  movel([-0.141321, -0.804315, -2.796072, -1.112001, 1.570796, 1.429476],accel_mss,speed_ms,0,blend_radius_m)
  movel([-0.146733, -0.812986, -2.794574, -1.104829, 1.570796, 1.424064],accel_mss,speed_ms,0,blend_radius_m)
  movel([-0.151447, -0.821414, -2.793080, -1.097895, 1.570796, 1.419350],accel_mss,speed_ms,0,blend_radius_m)
  movel([-0.155435, -0.829598, -2.791592, -1.091199, 1.570796, 1.415362],accel_mss,speed_ms,0,blend_radius_m)
  movel([-0.157149, -0.833600, -2.790851, -1.087938, 1.570796, 1.413648],accel_mss,speed_ms,0,blend_radius_m)
  movel([-0.159989, -0.841407, -2.789381, -1.081601, 1.570796, 1.410807],accel_mss,speed_ms,0,blend_radius_m)
  movel([-0.161109, -0.845218, -2.788651, -1.078520, 1.570796, 1.409688],accel_mss,speed_ms,0,blend_radius_m)
  movel([-0.162732, -0.852643, -2.787205, -1.072541, 1.570796, 1.408064],accel_mss,speed_ms,0,blend_radius_m)
  movel([-0.163230, -0.856264, -2.786488, -1.069637, 1.570796, 1.407566],accel_mss,speed_ms,0,blend_radius_m)
  movel([-0.163513, -0.859817, -2.785778, -1.066794, 1.570796, 1.407283],accel_mss,speed_ms,0,blend_radius_m)
  movel([-0.163602, -0.864722, -2.784786, -1.062881, 1.570796, 1.407194],accel_mss,speed_ms,0,blend_radius_m)
  movel([-0.163380, -0.869441, -2.783818, -1.059131, 1.570796, 1.407417],accel_mss,speed_ms,0,blend_radius_m)
  movel([-0.162870, -0.873957, -2.782879, -1.055553, 1.570796, 1.407926],accel_mss,speed_ms,0,blend_radius_m)
  movel([-0.162104, -0.878276, -2.781970, -1.052143, 1.570796, 1.408692],accel_mss,speed_ms,0,blend_radius_m)
  movel([-0.161097, -0.882370, -2.781098, -1.048921, 1.570796, 1.409700],accel_mss,speed_ms,0,blend_radius_m)
  movel([-0.159870, -0.886230, -2.780267, -1.045892, 1.570796, 1.410927],accel_mss,speed_ms,0,blend_radius_m)
  movel([-0.158448, -0.889851, -2.779479, -1.043059, 1.570796, 1.412348],accel_mss,speed_ms,0,blend_radius_m)
  movel([-0.156848, -0.893214, -2.778740, -1.040435, 1.570796, 1.413948],accel_mss,speed_ms,0,blend_radius_m)
  movel([-0.149158, -0.904985, -2.776098, -1.031305, 1.570796, 1.421638],accel_mss,speed_ms,0,blend_radius_m)
  movel([-0.143209, -0.914586, -2.773880, -1.023923, 1.570796, 1.427587],accel_mss,speed_ms,0,blend_radius_m)
  movel([-0.142775, -0.915615, -2.773639, -1.023135, 1.570796, 1.428021],accel_mss,speed_ms,0,blend_radius_m)
  movel([-0.135600, -0.906199, -2.775821, -1.030369, 1.570796, 1.435197],accel_mss,speed_ms,0,blend_radius_m)
  movel([-0.127938, -0.896903, -2.777921, -1.037564, 1.570796, 1.442859],accel_mss,speed_ms,0,blend_radius_m)
  movel([-0.119839, -0.887763, -2.779934, -1.044692, 1.570796, 1.450957],accel_mss,speed_ms,0,blend_radius_m)
  movel([-0.111369, -0.878821, -2.781854, -1.051713, 1.570796, 1.459427],accel_mss,speed_ms,0,blend_radius_m)
  movel([-0.102591, -0.870130, -2.783675, -1.058584, 1.570796, 1.468205],accel_mss,speed_ms,0,blend_radius_m)
  movel([-0.093574, -0.861730, -2.785393, -1.065267, 1.570796, 1.477222],accel_mss,speed_ms,0,blend_radius_m)
  movel([-0.084386, -0.853674, -2.787002, -1.071713, 1.570796, 1.486410],accel_mss,speed_ms,0,blend_radius_m)
  movel([-0.075105, -0.846013, -2.788497, -1.077879, 1.570796, 1.495692],accel_mss,speed_ms,0,blend_radius_m)
  movel([-0.070692, -0.842600, -2.789153, -1.080635, 1.570796, 1.500104],accel_mss,speed_ms,0,blend_radius_m)
  movel([-0.066171, -0.839349, -2.789772, -1.083268, 1.570796, 1.504626],accel_mss,speed_ms,0,blend_radius_m)
  movel([-0.061579, -0.836295, -2.790347, -1.085746, 1.570796, 1.509218],accel_mss,speed_ms,0,blend_radius_m)
  movel([-0.056967, -0.833486, -2.790873, -1.088031, 1.570796, 1.513830],accel_mss,speed_ms,0,blend_radius_m)
  movel([-0.052375, -0.830958, -2.791341, -1.090090, 1.570796, 1.518421],accel_mss,speed_ms,0,blend_radius_m)
  movel([-0.047846, -0.828755, -2.791747, -1.091887, 1.570796, 1.522951],accel_mss,speed_ms,0,blend_radius_m)
  movel([-0.043425, -0.826913, -2.792084, -1.093392, 1.570796, 1.527371],accel_mss,speed_ms,0,blend_radius_m)
  movel([-0.039161, -0.825474, -2.792346, -1.094569, 1.570796, 1.531636],accel_mss,speed_ms,0,blend_radius_m)
  movel([-0.035094, -0.824478, -2.792527, -1.095384, 1.570796, 1.535702],accel_mss,speed_ms,0,blend_radius_m)
  movel([-0.031268, -0.823960, -2.792621, -1.095808, 1.570796, 1.539528],accel_mss,speed_ms,0,blend_radius_m)
  movel([-0.027734, -0.823963, -2.792620, -1.095806, 1.570796, 1.543062],accel_mss,speed_ms,0,blend_radius_m)
  movel([-0.024533, -0.824519, -2.792520, -1.095350, 1.570796, 1.546264],accel_mss,speed_ms,0,blend_radius_m)
  movel([-0.021709, -0.825663, -2.792312, -1.094414, 1.570796, 1.549087],accel_mss,speed_ms,0,blend_radius_m)
  movel([-0.019297, -0.827423, -2.791991, -1.092975, 1.570796, 1.551499],accel_mss,speed_ms,0,blend_radius_m)
  movel([-0.017345, -0.829831, -2.791549, -1.091009, 1.570796, 1.553452],accel_mss,speed_ms,0,blend_radius_m)
  movel([-0.015891, -0.832916, -2.790978, -1.088494, 1.570796, 1.554905],accel_mss,speed_ms,0,blend_radius_m)
  movel([-0.014708, -0.837711, -2.790081, -1.084597, 1.570796, 1.556088],accel_mss,speed_ms,0,blend_radius_m)
  movel([-0.014174, -0.843160, -2.789046, -1.080183, 1.570796, 1.556622],accel_mss,speed_ms,0,blend_radius_m)
  movel([-0.014196, -0.849111, -2.787897, -1.075382, 1.570796, 1.556600],accel_mss,speed_ms,0,blend_radius_m)
  movel([-0.014673, -0.855417, -2.786657, -1.070315, 1.570796, 1.556123],accel_mss,speed_ms,0,blend_radius_m)
  movel([-0.015515, -0.861935, -2.785351, -1.065103, 1.570796, 1.555282],accel_mss,speed_ms,0,blend_radius_m)
  movel([-0.016634, -0.868531, -2.784005, -1.059853, 1.570796, 1.554162],accel_mss,speed_ms,0,blend_radius_m)
  movel([-0.019330, -0.881416, -2.781302, -1.049671, 1.570796, 1.551466],accel_mss,speed_ms,0,blend_radius_m)
  movel([-0.021385, -0.889588, -2.779536, -1.043265, 1.570796, 1.549411],accel_mss,speed_ms,0,blend_radius_m)
  movel([-0.023782, -0.897714, -2.777740, -1.036935, 1.570796, 1.547015],accel_mss,speed_ms,0,blend_radius_m)
  movel([-0.026474, -0.905794, -2.775914, -1.030681, 1.570796, 1.544323],accel_mss,speed_ms,0,blend_radius_m)
  movel([-0.029419, -0.913847, -2.774053, -1.024489, 1.570796, 1.541377],accel_mss,speed_ms,0,blend_radius_m)
  movel([-0.032573, -0.921870, -2.772158, -1.018361, 1.570796, 1.538223],accel_mss,speed_ms,0,blend_radius_m)
  movel([-0.035892, -0.929878, -2.770225, -1.012287, 1.570796, 1.534904],accel_mss,speed_ms,0,blend_radius_m)
  movel([-0.042880, -0.945892, -2.766232, -1.000265, 1.570796, 1.527916],accel_mss,speed_ms,0,blend_radius_m)
  movel([-0.036325, -0.946186, -2.766157, -1.000046, 1.570796, 1.534471],accel_mss,speed_ms,0,blend_radius_m)
  movel([-0.032953, -0.946594, -2.766053, -0.999742, 1.570796, 1.537843],accel_mss,speed_ms,0,blend_radius_m)
  movel([-0.030089, -0.947502, -2.765821, -0.999065, 1.570796, 1.540707],accel_mss,speed_ms,0,blend_radius_m)
  movel([-0.028984, -0.948223, -2.765637, -0.998529, 1.570796, 1.541813],accel_mss,speed_ms,0,blend_radius_m)
  movel([-0.028168, -0.949162, -2.765396, -0.997831, 1.570796, 1.542628],accel_mss,speed_ms,0,blend_radius_m)
  movel([-0.027690, -0.950344, -2.765092, -0.996953, 1.570796, 1.543106],accel_mss,speed_ms,0,blend_radius_m)
  movel([-0.027603, -0.951798, -2.764716, -0.995875, 1.570796, 1.543193],accel_mss,speed_ms,0,blend_radius_m)
  movel([-0.027958, -0.953548, -2.764263, -0.994579, 1.570796, 1.542838],accel_mss,speed_ms,0,blend_radius_m)
  movel([-0.028810, -0.955631, -2.763720, -0.993039, 1.570796, 1.541986],accel_mss,speed_ms,0,blend_radius_m)
  movel([-0.030204, -0.958070, -2.763080, -0.991239, 1.570796, 1.540592],accel_mss,speed_ms,0,blend_radius_m)
  movel([-0.032189, -0.960886, -2.762337, -0.989166, 1.570796, 1.538607],accel_mss,speed_ms,0,blend_radius_m)
  movel([-0.034030, -0.963178, -2.761728, -0.987484, 1.570796, 1.536766],accel_mss,speed_ms,0,blend_radius_m)
  movel([-0.035882, -0.965239, -2.761177, -0.985973, 1.570796, 1.534914],accel_mss,speed_ms,0,blend_radius_m)
  movel([-0.037742, -0.967088, -2.760680, -0.984621, 1.570796, 1.533055],accel_mss,speed_ms,0,blend_radius_m)
  movel([-0.041487, -0.970225, -2.759832, -0.982332, 1.570796, 1.529310],accel_mss,speed_ms,0,blend_radius_m)
  movel([-0.043369, -0.971550, -2.759471, -0.981368, 1.570796, 1.527427],accel_mss,speed_ms,0,blend_radius_m)
  movel([-0.047159, -0.973809, -2.758854, -0.979726, 1.570796, 1.523638],accel_mss,speed_ms,0,blend_radius_m)
  movel([-0.050963, -0.975658, -2.758346, -0.978385, 1.570796, 1.519833],accel_mss,speed_ms,0,blend_radius_m)
  movel([-0.054779, -0.977239, -2.757910, -0.977241, 1.570796, 1.516017],accel_mss,speed_ms,0,blend_radius_m)
  movel([-0.062394, -0.980130, -2.757107, -0.975152, 1.570796, 1.508402],accel_mss,speed_ms,0,blend_radius_m)
  movel([-0.066370, -0.986523, -2.755311, -0.970555, 1.570796, 1.504426],accel_mss,speed_ms,0,blend_radius_m)
  movel([-0.068546, -0.989715, -2.754403, -0.968271, 1.570796, 1.502250],accel_mss,speed_ms,0,blend_radius_m)
  movel([-0.070857, -0.992817, -2.753513, -0.966058, 1.570796, 1.499939],accel_mss,speed_ms,0,blend_radius_m)
  movel([-0.073309, -0.995761, -2.752662, -0.963965, 1.570796, 1.497488],accel_mss,speed_ms,0,blend_radius_m)
  movel([-0.075903, -0.998481, -2.751871, -0.962038, 1.570796, 1.494894],accel_mss,speed_ms,0,blend_radius_m)
  movel([-0.078648, -1.000910, -2.751159, -0.960321, 1.570796, 1.492149],accel_mss,speed_ms,0,blend_radius_m)
  movel([-0.081555, -1.002990, -2.750546, -0.958854, 1.570796, 1.489241],accel_mss,speed_ms,0,blend_radius_m)
  movel([-0.083598, -1.004037, -2.750236, -0.958116, 1.570796, 1.487198],accel_mss,speed_ms,0,blend_radius_m)
  movel([-0.085214, -1.004394, -2.750130, -0.957865, 1.570796, 1.485582],accel_mss,speed_ms,0,blend_radius_m)
  movel([-0.086450, -1.004162, -2.750199, -0.958028, 1.570796, 1.484347],accel_mss,speed_ms,0,blend_radius_m)
  movel([-0.087346, -1.003436, -2.750414, -0.958539, 1.570796, 1.483451],accel_mss,speed_ms,0,blend_radius_m)
  movel([-0.087946, -1.002312, -2.750746, -0.959331, 1.570796, 1.482851],accel_mss,speed_ms,0,blend_radius_m)
  movel([-0.088287, -1.000895, -2.751163, -0.960331, 1.570796, 1.482509],accel_mss,speed_ms,0,blend_radius_m)
  movel([-0.088418, -0.999280, -2.751637, -0.961472, 1.570796, 1.482378],accel_mss,speed_ms,0,blend_radius_m)
  movel([-0.088369, -0.997561, -2.752139, -0.962689, 1.570796, 1.482428],accel_mss,speed_ms,0,blend_radius_m)
  movel([-0.087893, -0.993747, -2.753245, -0.965397, 1.570796, 1.482904],accel_mss,speed_ms,0,blend_radius_m)
  movel([-0.087059, -0.989798, -2.754379, -0.968212, 1.570796, 1.483737],accel_mss,speed_ms,0,blend_radius_m)
  movel([-0.084858, -0.981561, -2.756707, -0.974120, 1.570796, 1.485939],accel_mss,speed_ms,0,blend_radius_m)
  movel([-0.093540, -0.980140, -2.757104, -0.975145, 1.570796, 1.477256],accel_mss,speed_ms,0,blend_radius_m)
  movel([-0.102455, -0.979099, -2.757394, -0.975896, 1.570796, 1.468341],accel_mss,speed_ms,0,blend_radius_m)
  movel([-0.111365, -0.978026, -2.757692, -0.976671, 1.570796, 1.459431],accel_mss,speed_ms,0,blend_radius_m)
  movel([-0.115747, -0.977350, -2.757879, -0.977161, 1.570796, 1.455049],accel_mss,speed_ms,0,blend_radius_m)
  movel([-0.120046, -0.976509, -2.758111, -0.977769, 1.570796, 1.450750],accel_mss,speed_ms,0,blend_radius_m)
  movel([-0.124039, -0.975495, -2.758391, -0.978503, 1.570796, 1.446757],accel_mss,speed_ms,0,blend_radius_m)
  movel([-0.127889, -0.974301, -2.758719, -0.979369, 1.570796, 1.442907],accel_mss,speed_ms,0,blend_radius_m)
  movel([-0.135327, -0.971570, -2.759466, -0.981353, 1.570796, 1.435469],accel_mss,speed_ms,0,blend_radius_m)
  movel([-0.142709, -0.968772, -2.760225, -0.983392, 1.570796, 1.428087],accel_mss,speed_ms,0,blend_radius_m)
  movel([-0.150371, -0.966361, -2.760875, -0.985152, 1.570796, 1.420425],accel_mss,speed_ms,0,blend_radius_m)
  movel([-0.152086, -0.971127, -2.759586, -0.981675, 1.570796, 1.418710],accel_mss,speed_ms,0,blend_radius_m)
  movel([-0.153549, -0.975769, -2.758315, -0.978305, 1.570796, 1.417247],accel_mss,speed_ms,0,blend_radius_m)
  movel([-0.154762, -0.980277, -2.757066, -0.975046, 1.570796, 1.416035],accel_mss,speed_ms,0,blend_radius_m)
  movel([-0.155729, -0.984644, -2.755842, -0.971903, 1.570796, 1.415067],accel_mss,speed_ms,0,blend_radius_m)
  movel([-0.156451, -0.988870, -2.754644, -0.968875, 1.570796, 1.414345],accel_mss,speed_ms,0,blend_radius_m)
  movel([-0.156938, -0.992946, -2.753476, -0.965967, 1.570796, 1.413859],accel_mss,speed_ms,0,blend_radius_m)
  movel([-0.157185, -0.996868, -2.752341, -0.963180, 1.570796, 1.413612],accel_mss,speed_ms,0,blend_radius_m)
  movel([-0.157205, -1.000637, -2.751239, -0.960513, 1.570796, 1.413592],accel_mss,speed_ms,0,blend_radius_m)
  movel([-0.156995, -1.004243, -2.750175, -0.957972, 1.570796, 1.413802],accel_mss,speed_ms,0,blend_radius_m)
  movel([-0.156554, -1.007678, -2.749152, -0.955559, 1.570796, 1.414242],accel_mss,speed_ms,0,blend_radius_m)
  movel([-0.155895, -1.010950, -2.748169, -0.953270, 1.570796, 1.414901],accel_mss,speed_ms,0,blend_radius_m)
  movel([-0.155018, -1.014046, -2.747232, -0.951112, 1.570796, 1.415778],accel_mss,speed_ms,0,blend_radius_m)
  movel([-0.153919, -1.016958, -2.746343, -0.949088, 1.570796, 1.416877],accel_mss,speed_ms,0,blend_radius_m)
  movel([-0.152607, -1.019693, -2.745503, -0.947193, 1.570796, 1.418189],accel_mss,speed_ms,0,blend_radius_m)
  movel([-0.151084, -1.022240, -2.744715, -0.945434, 1.570796, 1.419713],accel_mss,speed_ms,0,blend_radius_m)
  movel([-0.149346, -1.024596, -2.743981, -0.943812, 1.570796, 1.421450],accel_mss,speed_ms,0,blend_radius_m)
  movel([-0.146282, -1.027856, -2.742959, -0.941574, 1.570796, 1.424514],accel_mss,speed_ms,0,blend_radius_m)
  movel([-0.142850, -1.030642, -2.742079, -0.939668, 1.570796, 1.427946],accel_mss,speed_ms,0,blend_radius_m)
  movel([-0.139097, -1.033005, -2.741328, -0.938057, 1.570796, 1.431699],accel_mss,speed_ms,0,blend_radius_m)
  movel([-0.135055, -1.034984, -2.740695, -0.936710, 1.570796, 1.435741],accel_mss,speed_ms,0,blend_radius_m)
  movel([-0.130770, -1.036629, -2.740167, -0.935593, 1.570796, 1.440026],accel_mss,speed_ms,0,blend_radius_m)
  movel([-0.126280, -1.037978, -2.739732, -0.934679, 1.570796, 1.444516],accel_mss,speed_ms,0,blend_radius_m)
  movel([-0.121626, -1.039078, -2.739376, -0.933935, 1.570796, 1.449171],accel_mss,speed_ms,0,blend_radius_m)
  movel([-0.116838, -1.039956, -2.739092, -0.933342, 1.570796, 1.453958],accel_mss,speed_ms,0,blend_radius_m)
  movel([-0.106974, -1.041285, -2.738660, -0.932445, 1.570796, 1.463822],accel_mss,speed_ms,0,blend_radius_m)
  movel([-0.096981, -1.042372, -2.738305, -0.931712, 1.570796, 1.473815],accel_mss,speed_ms,0,blend_radius_m)
  movel([-0.089406, -1.043472, -2.737946, -0.930972, 1.570796, 1.481391],accel_mss,speed_ms,0,blend_radius_m)
  movel([-0.086797, -1.043644, -2.737889, -0.930856, 1.570796, 1.484000],accel_mss,speed_ms,0,blend_radius_m)
  movel([-0.082087, -1.043552, -2.737919, -0.930918, 1.570796, 1.488709],accel_mss,speed_ms,0,blend_radius_m)
  movel([-0.081105, -1.043729, -2.737861, -0.930799, 1.570796, 1.489692],accel_mss,speed_ms,0,blend_radius_m)
  movel([-0.080223, -1.044102, -2.737739, -0.930548, 1.570796, 1.490574],accel_mss,speed_ms,0,blend_radius_m)
  movel([-0.079458, -1.044736, -2.737531, -0.930122, 1.570796, 1.491338],accel_mss,speed_ms,0,blend_radius_m)
  movel([-0.078830, -1.045693, -2.737216, -0.929480, 1.570796, 1.491966],accel_mss,speed_ms,0,blend_radius_m)
  movel([-0.078371, -1.047037, -2.736773, -0.928579, 1.570796, 1.492426],accel_mss,speed_ms,0,blend_radius_m)
  movel([-0.078211, -1.048560, -2.736269, -0.927560, 1.570796, 1.492585],accel_mss,speed_ms,0,blend_radius_m)
  movel([-0.078322, -1.050228, -2.735715, -0.926446, 1.570796, 1.492474],accel_mss,speed_ms,0,blend_radius_m)
  movel([-0.078680, -1.052026, -2.735115, -0.925248, 1.570796, 1.492116],accel_mss,speed_ms,0,blend_radius_m)
  movel([-0.079260, -1.053920, -2.734480, -0.923989, 1.570796, 1.491536],accel_mss,speed_ms,0,blend_radius_m)
  movel([-0.080989, -1.057919, -2.733129, -0.921340, 1.570796, 1.489808],accel_mss,speed_ms,0,blend_radius_m)
  movel([-0.082090, -1.059975, -2.732430, -0.919984, 1.570796, 1.488706],accel_mss,speed_ms,0,blend_radius_m)
  movel([-0.084632, -1.064080, -2.731023, -0.917287, 1.570796, 1.486165],accel_mss,speed_ms,0,blend_radius_m)
  movel([-0.087485, -1.068033, -2.729654, -0.914703, 1.570796, 1.483311],accel_mss,speed_ms,0,blend_radius_m)
  movel([-0.090454, -1.071655, -2.728388, -0.912347, 1.570796, 1.480342],accel_mss,speed_ms,0,blend_radius_m)
  movel([-0.093367, -1.074779, -2.727286, -0.910323, 1.570796, 1.477429],accel_mss,speed_ms,0,blend_radius_m)
  movel([-0.097927, -1.079003, -2.725784, -0.907602, 1.570796, 1.472870],accel_mss,speed_ms,0,blend_radius_m)
  movel([-0.100289, -1.080959, -2.725083, -0.906347, 1.570796, 1.470507],accel_mss,speed_ms,0,blend_radius_m)
  movel([-0.102689, -1.082800, -2.724421, -0.905168, 1.570796, 1.468107],accel_mss,speed_ms,0,blend_radius_m)
  movel([-0.107574, -1.086135, -2.723212, -0.903042, 1.570796, 1.463222],accel_mss,speed_ms,0,blend_radius_m)
  movel([-0.112504, -1.088976, -2.722175, -0.901238, 1.570796, 1.458292],accel_mss,speed_ms,0,blend_radius_m)
  movel([-0.117406, -1.091288, -2.721326, -0.899775, 1.570796, 1.453391],accel_mss,speed_ms,0,blend_radius_m)
  movel([-0.122195, -1.093035, -2.720681, -0.898673, 1.570796, 1.448602],accel_mss,speed_ms,0,blend_radius_m)
  movel([-0.124527, -1.093683, -2.720441, -0.898265, 1.570796, 1.446270],accel_mss,speed_ms,0,blend_radius_m)
  movel([-0.129018, -1.094511, -2.720134, -0.897744, 1.570796, 1.441778],accel_mss,speed_ms,0,blend_radius_m)
  movel([-0.131158, -1.094678, -2.720072, -0.897639, 1.570796, 1.439638],accel_mss,speed_ms,0,blend_radius_m)
  movel([-0.133875, -1.094654, -2.720081, -0.897654, 1.570796, 1.436921],accel_mss,speed_ms,0,blend_radius_m)
  movel([-0.136457, -1.094390, -2.720179, -0.897821, 1.570796, 1.434339],accel_mss,speed_ms,0,blend_radius_m)
  movel([-0.138916, -1.093913, -2.720356, -0.898121, 1.570796, 1.431880],accel_mss,speed_ms,0,blend_radius_m)
  movel([-0.141274, -1.093262, -2.720597, -0.898530, 1.570796, 1.429522],accel_mss,speed_ms,0,blend_radius_m)
  movel([-0.145748, -1.091559, -2.721226, -0.899604, 1.570796, 1.425048],accel_mss,speed_ms,0,blend_radius_m)
  movel([-0.150009, -1.089547, -2.721966, -0.900876, 1.570796, 1.420787],accel_mss,speed_ms,0,blend_radius_m)
  movel([-0.155186, -1.086801, -2.722970, -0.902618, 1.570796, 1.415610],accel_mss,speed_ms,0,blend_radius_m)
  movel([-0.160187, -1.083750, -2.724077, -0.904561, 1.570796, 1.410610],accel_mss,speed_ms,0,blend_radius_m)
  movel([-0.164967, -1.080374, -2.725293, -0.906722, 1.570796, 1.405830],accel_mss,speed_ms,0,blend_radius_m)
  movel([-0.169489, -1.076653, -2.726622, -0.909114, 1.570796, 1.401308],accel_mss,speed_ms,0,blend_radius_m)
  movel([-0.173708, -1.072561, -2.728069, -0.911759, 1.570796, 1.397089],accel_mss,speed_ms,0,blend_radius_m)
  movel([-0.177576, -1.068074, -2.729639, -0.914676, 1.570796, 1.393221],accel_mss,speed_ms,0,blend_radius_m)
  movel([-0.181051, -1.063167, -2.731337, -0.917886, 1.570796, 1.389745],accel_mss,speed_ms,0,blend_radius_m)
  movel([-0.184087, -1.057810, -2.733166, -0.921412, 1.570796, 1.386710],accel_mss,speed_ms,0,blend_radius_m)
  movel([-0.186073, -1.053486, -2.734626, -0.924278, 1.570796, 1.384723],accel_mss,speed_ms,0,blend_radius_m)
  movel([-0.187880, -1.048763, -2.736202, -0.927424, 1.570796, 1.382916],accel_mss,speed_ms,0,blend_radius_m)
  movel([-0.189439, -1.043669, -2.737881, -0.930839, 1.570796, 1.381358],accel_mss,speed_ms,0,blend_radius_m)
  movel([-0.190682, -1.038239, -2.739647, -0.934502, 1.570796, 1.380114],accel_mss,speed_ms,0,blend_radius_m)
  movel([-0.191534, -1.032503, -2.741488, -0.938398, 1.570796, 1.379263],accel_mss,speed_ms,0,blend_radius_m)
  movel([-0.191918, -1.026493, -2.743388, -0.942509, 1.570796, 1.378878],accel_mss,speed_ms,0,blend_radius_m)
  movel([-0.191763, -1.020236, -2.745335, -0.946818, 1.570796, 1.379033],accel_mss,speed_ms,0,blend_radius_m)
  movel([-0.191455, -1.017023, -2.746323, -0.949042, 1.570796, 1.379341],accel_mss,speed_ms,0,blend_radius_m)
  movel([-0.190983, -1.013763, -2.747318, -0.951308, 1.570796, 1.379813],accel_mss,speed_ms,0,blend_radius_m)
  movel([-0.189719, -1.007476, -2.749212, -0.955701, 1.570796, 1.381077],accel_mss,speed_ms,0,blend_radius_m)
  movel([-0.188031, -1.000973, -2.751140, -0.960275, 1.570796, 1.382765],accel_mss,speed_ms,0,blend_radius_m)
  movel([-0.185918, -0.994276, -2.753093, -0.965021, 1.570796, 1.384878],accel_mss,speed_ms,0,blend_radius_m)
  movel([-0.183392, -0.987409, -2.755060, -0.969921, 1.570796, 1.387404],accel_mss,speed_ms,0,blend_radius_m)
  movel([-0.180442, -0.980392, -2.757034, -0.974963, 1.570796, 1.390354],accel_mss,speed_ms,0,blend_radius_m)
  movel([-0.177085, -0.973259, -2.759004, -0.980126, 1.570796, 1.393711],accel_mss,speed_ms,0,blend_radius_m)
  movel([-0.173317, -0.966031, -2.760964, -0.985394, 1.570796, 1.397479],accel_mss,speed_ms,0,blend_radius_m)
  movel([-0.169142, -0.958742, -2.762903, -0.990744, 1.570796, 1.401654],accel_mss,speed_ms,0,blend_radius_m)
  movel([-0.177984, -0.951083, -2.764901, -0.996405, 1.570796, 1.392812],accel_mss,speed_ms,0,blend_radius_m)
  movel([-0.182461, -0.947285, -2.765877, -0.999227, 1.570796, 1.388335],accel_mss,speed_ms,0,blend_radius_m)
  movel([-0.186722, -0.943199, -2.766916, -1.002275, 1.570796, 1.384074],accel_mss,speed_ms,0,blend_radius_m)
  movel([-0.189559, -0.939742, -2.767786, -1.004861, 1.570796, 1.381237],accel_mss,speed_ms,0,blend_radius_m)
  movel([-0.191976, -0.935811, -2.768765, -1.007813, 1.570796, 1.378820],accel_mss,speed_ms,0,blend_radius_m)
  movel([-0.193988, -0.931437, -2.769843, -1.011108, 1.570796, 1.376808],accel_mss,speed_ms,0,blend_radius_m)
  movel([-0.195602, -0.926639, -2.771012, -1.014739, 1.570796, 1.375194],accel_mss,speed_ms,0,blend_radius_m)
  movel([-0.196828, -0.921444, -2.772259, -1.018685, 1.570796, 1.373968],accel_mss,speed_ms,0,blend_radius_m)
  movel([-0.197671, -0.915875, -2.773578, -1.022936, 1.570796, 1.373125],accel_mss,speed_ms,0,blend_radius_m)
  movel([-0.198141, -0.909954, -2.774958, -1.027477, 1.570796, 1.372655],accel_mss,speed_ms,0,blend_radius_m)
  movel([-0.198246, -0.903710, -2.776389, -1.032290, 1.570796, 1.372550],accel_mss,speed_ms,0,blend_radius_m)
  movel([-0.197990, -0.897171, -2.777862, -1.037356, 1.570796, 1.372806],accel_mss,speed_ms,0,blend_radius_m)
  movel([-0.197379, -0.890353, -2.779369, -1.042667, 1.570796, 1.373418],accel_mss,speed_ms,0,blend_radius_m)
  movel([-0.196419, -0.883290, -2.780901, -1.048198, 1.570796, 1.374377],accel_mss,speed_ms,0,blend_radius_m)
  movel([-0.195120, -0.876011, -2.782448, -1.053930, 1.570796, 1.375676],accel_mss,speed_ms,0,blend_radius_m)
  movel([-0.193486, -0.868544, -2.784003, -1.059842, 1.570796, 1.377310],accel_mss,speed_ms,0,blend_radius_m)
  movel([-0.191530, -0.860930, -2.785554, -1.065905, 1.570796, 1.379267],accel_mss,speed_ms,0,blend_radius_m)
  movel([-0.189249, -0.853187, -2.787098, -1.072104, 1.570796, 1.381547],accel_mss,speed_ms,0,blend_radius_m)
  movel([-0.186663, -0.845361, -2.788623, -1.078405, 1.570796, 1.384133],accel_mss,speed_ms,0,blend_radius_m)
  movel([-0.181160, -0.830361, -2.791451, -1.090576, 1.570796, 1.389637],accel_mss,speed_ms,0,blend_radius_m)
  movel([-0.178053, -0.822646, -2.792858, -1.096885, 1.570796, 1.392744],accel_mss,speed_ms,0,blend_radius_m)
  movel([-0.174652, -0.814792, -2.794257, -1.103340, 1.570796, 1.396144],accel_mss,speed_ms,0,blend_radius_m)
  movel([-0.170903, -0.806807, -2.795646, -1.109936, 1.570796, 1.399893],accel_mss,speed_ms,0,blend_radius_m)
  movel([-0.166766, -0.798708, -2.797020, -1.116660, 1.570796, 1.404030],accel_mss,speed_ms,0,blend_radius_m)
  movel([-0.162191, -0.790498, -2.798379, -1.123512, 1.570796, 1.408605],accel_mss,speed_ms,0,blend_radius_m)
  movel([-0.157128, -0.782189, -2.799719, -1.130481, 1.570796, 1.413668],accel_mss,speed_ms,0,blend_radius_m)
  movel([-0.150973, -0.772894, -2.801177, -1.138318, 1.570796, 1.419823],accel_mss,speed_ms,0,blend_radius_m)
  movel([-0.144342, -0.763571, -2.802597, -1.146221, 1.570796, 1.426454],accel_mss,speed_ms,0,blend_radius_m)
  movel([-0.137271, -0.754250, -2.803974, -1.154165, 1.570796, 1.433525],accel_mss,speed_ms,0,blend_radius_m)
  movel([-0.129792, -0.744968, -2.805304, -1.162117, 1.570796, 1.441004],accel_mss,speed_ms,0,blend_radius_m)
  movel([-0.121944, -0.735767, -2.806582, -1.170041, 1.570796, 1.448852],accel_mss,speed_ms,0,blend_radius_m)
  movel([-0.113770, -0.726690, -2.807804, -1.177895, 1.570796, 1.457026],accel_mss,speed_ms,0,blend_radius_m)
  movel([-0.105305, -0.717773, -2.808968, -1.185648, 1.570796, 1.465492],accel_mss,speed_ms,0,blend_radius_m)
  movel([-0.096600, -0.709069, -2.810069, -1.193251, 1.570796, 1.474197],accel_mss,speed_ms,0,blend_radius_m)
  movel([-0.087699, -0.700626, -2.811105, -1.200658, 1.570796, 1.483097],accel_mss,speed_ms,0,blend_radius_m)
  movel([-0.078662, -0.692490, -2.812073, -1.207826, 1.570796, 1.492134],accel_mss,speed_ms,0,blend_radius_m)
  movel([-0.069532, -0.684712, -2.812972, -1.214705, 1.570796, 1.501264],accel_mss,speed_ms,0,blend_radius_m)
  movel([-0.060365, -0.677340, -2.813799, -1.221250, 1.570796, 1.510431],accel_mss,speed_ms,0,blend_radius_m)
  movel([-0.051227, -0.670430, -2.814554, -1.227404, 1.570796, 1.519569],accel_mss,speed_ms,0,blend_radius_m)
  movel([-0.042167, -0.664027, -2.815235, -1.233126, 1.570796, 1.528629],accel_mss,speed_ms,0,blend_radius_m)
  movel([-0.033247, -0.658183, -2.815842, -1.238364, 1.570796, 1.537549],accel_mss,speed_ms,0,blend_radius_m)
  movel([-0.024524, -0.652948, -2.816374, -1.243067, 1.570796, 1.546273],accel_mss,speed_ms,0,blend_radius_m)
  movel([-0.015396, -0.647880, -2.816878, -1.247631, 1.570796, 1.555400],accel_mss,speed_ms,0,blend_radius_m)
  movel([-0.006368, -0.643230, -2.817331, -1.251828, 1.570796, 1.564428],accel_mss,speed_ms,0,blend_radius_m)
  movel([0.002483, -0.639132, -2.817723, -1.255535, 1.570796, 1.573279],accel_mss,speed_ms,0,blend_radius_m)
  movel([0.011077, -0.635735, -2.818042, -1.258611, 1.570796, 1.581874],accel_mss,speed_ms,0,blend_radius_m)
  movel([0.020717, -0.632779, -2.818317, -1.261293, 1.570796, 1.591514],accel_mss,speed_ms,0,blend_radius_m)
  movel([0.029958, -0.630878, -2.818491, -1.263019, 1.570796, 1.600754],accel_mss,speed_ms,0,blend_radius_m)
  movel([0.038695, -0.630051, -2.818567, -1.263771, 1.570796, 1.609491],accel_mss,speed_ms,0,blend_radius_m)
  movel([0.046827, -0.630306, -2.818544, -1.263539, 1.570796, 1.617623],accel_mss,speed_ms,0,blend_radius_m)
  movel([0.054267, -0.631639, -2.818422, -1.262328, 1.570796, 1.625063],accel_mss,speed_ms,0,blend_radius_m)
  movel([0.060928, -0.634042, -2.818200, -1.260147, 1.570796, 1.631725],accel_mss,speed_ms,0,blend_radius_m)
  movel([0.066738, -0.637486, -2.817878, -1.257025, 1.570796, 1.637535],accel_mss,speed_ms,0,blend_radius_m)
  movel([0.071630, -0.641948, -2.817454, -1.252987, 1.570796, 1.642427],accel_mss,speed_ms,0,blend_radius_m)
  movel([0.080139, -0.652079, -2.816461, -1.243849, 1.570796, 1.650935],accel_mss,speed_ms,0,blend_radius_m)
  movel([0.083892, -0.657646, -2.815897, -1.238846, 1.570796, 1.654688],accel_mss,speed_ms,0,blend_radius_m)
  movel([0.087126, -0.663924, -2.815246, -1.233219, 1.570796, 1.657922],accel_mss,speed_ms,0,blend_radius_m)
  movel([0.092254, -0.674828, -2.814076, -1.223485, 1.570796, 1.663050],accel_mss,speed_ms,0,blend_radius_m)
  movel([0.095202, -0.679953, -2.813509, -1.218927, 1.570796, 1.665998],accel_mss,speed_ms,0,blend_radius_m)
  movel([0.098521, -0.684636, -2.812980, -1.214773, 1.570796, 1.669318],accel_mss,speed_ms,0,blend_radius_m)
  movel([0.102318, -0.688705, -2.812514, -1.211170, 1.570796, 1.673114],accel_mss,speed_ms,0,blend_radius_m)
  movel([0.106666, -0.692002, -2.812130, -1.208257, 1.570796, 1.677463],accel_mss,speed_ms,0,blend_radius_m)
  movel([0.111676, -0.694361, -2.811853, -1.206175, 1.570796, 1.682472],accel_mss,speed_ms,0,blend_radius_m)
  movel([0.117434, -0.695618, -2.811704, -1.205067, 1.570796, 1.688231],accel_mss,speed_ms,0,blend_radius_m)
  movel([0.120030, -0.695672, -2.811698, -1.205019, 1.570796, 1.690827],accel_mss,speed_ms,0,blend_radius_m)
  movel([0.122938, -0.695135, -2.811761, -1.205492, 1.570796, 1.693735],accel_mss,speed_ms,0,blend_radius_m)
  movel([0.124501, -0.694553, -2.811830, -1.206006, 1.570796, 1.695297],accel_mss,speed_ms,0,blend_radius_m)
  movel([0.126126, -0.693719, -2.811928, -1.206741, 1.570796, 1.696922],accel_mss,speed_ms,0,blend_radius_m)
  movel([0.127815, -0.692594, -2.812061, -1.207734, 1.570796, 1.698611],accel_mss,speed_ms,0,blend_radius_m)
  movel([0.129555, -0.691139, -2.812231, -1.209019, 1.570796, 1.700351],accel_mss,speed_ms,0,blend_radius_m)
  movel([0.131319, -0.689354, -2.812438, -1.210597, 1.570796, 1.702115],accel_mss,speed_ms,0,blend_radius_m)
  movel([0.132980, -0.687374, -2.812667, -1.212348, 1.570796, 1.703776],accel_mss,speed_ms,0,blend_radius_m)
  movel([0.135970, -0.683096, -2.813155, -1.216138, 1.570796, 1.706767],accel_mss,speed_ms,0,blend_radius_m)
  movel([0.137783, -0.680045, -2.813498, -1.218845, 1.570796, 1.708580],accel_mss,speed_ms,0,blend_radius_m)
  movel([0.139361, -0.677032, -2.813833, -1.221523, 1.570796, 1.710157],accel_mss,speed_ms,0,blend_radius_m)
  movel([0.141870, -0.671141, -2.814477, -1.226770, 1.570796, 1.712666],accel_mss,speed_ms,0,blend_radius_m)
  movel([0.143598, -0.665477, -2.815083, -1.231830, 1.570796, 1.714394],accel_mss,speed_ms,0,blend_radius_m)
  movel([0.144658, -0.660075, -2.815647, -1.236667, 1.570796, 1.715454],accel_mss,speed_ms,0,blend_radius_m)
  movel([0.145152, -0.654997, -2.816167, -1.241224, 1.570796, 1.715948],accel_mss,speed_ms,0,blend_radius_m)
  movel([0.145192, -0.650285, -2.816640, -1.245464, 1.570796, 1.715988],accel_mss,speed_ms,0,blend_radius_m)
  movel([0.144887, -0.645985, -2.817063, -1.249341, 1.570796, 1.715683],accel_mss,speed_ms,0,blend_radius_m)
  movel([0.143440, -0.638102, -2.817820, -1.256467, 1.570796, 1.714237],accel_mss,speed_ms,0,blend_radius_m)
  movel([0.142144, -0.634435, -2.818164, -1.259791, 1.570796, 1.712941],accel_mss,speed_ms,0,blend_radius_m)
  movel([0.140471, -0.631159, -2.818466, -1.262764, 1.570796, 1.711267],accel_mss,speed_ms,0,blend_radius_m)
  movel([0.138417, -0.628311, -2.818725, -1.265353, 1.570796, 1.709214],accel_mss,speed_ms,0,blend_radius_m)
  movel([0.135985, -0.625905, -2.818941, -1.267543, 1.570796, 1.706781],accel_mss,speed_ms,0,blend_radius_m)
  movel([0.133177, -0.623970, -2.819114, -1.269305, 1.570796, 1.703974],accel_mss,speed_ms,0,blend_radius_m)
  movel([0.130010, -0.622516, -2.819242, -1.270631, 1.570796, 1.700806],accel_mss,speed_ms,0,blend_radius_m)
  movel([0.126480, -0.621568, -2.819326, -1.271496, 1.570796, 1.697276],accel_mss,speed_ms,0,blend_radius_m)
  speed_ms = 0.005
  movel([0.126480, -0.615674, -2.812529, -1.284186, 1.570796, 1.697276],accel_mss,speed_ms,0,blend_radius_m)
  speed_ms = 0.040
  movel([0.123325, -0.653236, -2.808959, -1.250194, 1.570796, 1.694121],accel_mss,speed_ms,0,blend_radius_m)
  speed_ms = 0.005
  movel([0.123325, -0.659726, -2.815683, -1.236980, 1.570796, 1.694121],accel_mss,speed_ms,0,blend_radius_m)
  speed_ms = 0.025
  movel([0.118895, -0.658973, -2.815761, -1.237654, 1.570796, 1.689691],accel_mss,speed_ms,0,blend_radius_m)
  movel([0.113905, -0.659116, -2.815746, -1.237527, 1.570796, 1.684701],accel_mss,speed_ms,0,blend_radius_m)
  movel([0.111148, -0.659712, -2.815685, -1.236992, 1.570796, 1.681944],accel_mss,speed_ms,0,blend_radius_m)
  movel([0.108196, -0.660754, -2.815577, -1.236058, 1.570796, 1.678993],accel_mss,speed_ms,0,blend_radius_m)
  movel([0.105036, -0.662312, -2.815415, -1.234662, 1.570796, 1.675833],accel_mss,speed_ms,0,blend_radius_m)
  movel([0.101649, -0.664453, -2.815191, -1.232745, 1.570796, 1.672446],accel_mss,speed_ms,0,blend_radius_m)
  speed_ms = 0.005
  movel([0.101649, -0.657892, -2.808476, -1.246022, 1.570796, 1.672446],accel_mss,speed_ms,0,blend_radius_m)
  speed_ms = 0.040
  movel([0.112275, -0.642742, -2.810015, -1.259632, 1.570796, 1.683072],accel_mss,speed_ms,0,blend_radius_m)
  speed_ms = 0.005
  movel([0.112275, -0.649070, -2.816760, -1.246559, 1.570796, 1.683072],accel_mss,speed_ms,0,blend_radius_m)
  speed_ms = 0.025
  movel([0.112399, -0.644194, -2.817238, -1.250958, 1.570796, 1.683195],accel_mss,speed_ms,0,blend_radius_m)
  movel([0.111517, -0.640308, -2.817611, -1.254471, 1.570796, 1.682314],accel_mss,speed_ms,0,blend_radius_m)
  movel([0.109701, -0.637442, -2.817882, -1.257065, 1.570796, 1.680497],accel_mss,speed_ms,0,blend_radius_m)
  movel([0.107011, -0.635659, -2.818049, -1.258681, 1.570796, 1.677807],accel_mss,speed_ms,0,blend_radius_m)
  movel([0.103521, -0.634994, -2.818111, -1.259283, 1.570796, 1.674318],accel_mss,speed_ms,0,blend_radius_m)
  movel([0.099319, -0.635483, -2.818066, -1.258840, 1.570796, 1.670115],accel_mss,speed_ms,0,blend_radius_m)
  movel([0.094491, -0.637147, -2.817910, -1.257332, 1.570796, 1.665287],accel_mss,speed_ms,0,blend_radius_m)
  movel([0.091867, -0.638433, -2.817789, -1.256167, 1.570796, 1.662663],accel_mss,speed_ms,0,blend_radius_m)
  movel([0.089124, -0.640011, -2.817639, -1.254739, 1.570796, 1.659920],accel_mss,speed_ms,0,blend_radius_m)
  speed_ms = 0.005
  movel([0.089124, -0.633823, -2.810876, -1.267689, 1.570796, 1.659920],accel_mss,speed_ms,0,blend_radius_m)
  speed_ms = 0.040
  movel([0.102652, -0.618294, -2.812299, -1.281796, 1.570796, 1.673448],accel_mss,speed_ms,0,blend_radius_m)
  speed_ms = 0.005
  movel([0.102652, -0.624231, -2.819091, -1.269067, 1.570796, 1.673448],accel_mss,speed_ms,0,blend_radius_m)
  speed_ms = 0.025
  movel([0.102279, -0.622165, -2.819273, -1.270951, 1.570796, 1.673075],accel_mss,speed_ms,0,blend_radius_m)
  movel([0.101580, -0.620373, -2.819430, -1.272586, 1.570796, 1.672376],accel_mss,speed_ms,0,blend_radius_m)
  movel([0.099284, -0.617623, -2.819669, -1.275097, 1.570796, 1.670080],accel_mss,speed_ms,0,blend_radius_m)
  movel([0.095934, -0.616002, -2.819808, -1.276579, 1.570796, 1.666730],accel_mss,speed_ms,0,blend_radius_m)
  movel([0.091712, -0.615526, -2.819849, -1.277014, 1.570796, 1.662509],accel_mss,speed_ms,0,blend_radius_m)
  movel([0.086803, -0.616184, -2.819792, -1.276413, 1.570796, 1.657599],accel_mss,speed_ms,0,blend_radius_m)
  movel([0.081418, -0.617958, -2.819640, -1.274791, 1.570796, 1.652214],accel_mss,speed_ms,0,blend_radius_m)
  movel([0.078603, -0.619264, -2.819527, -1.273598, 1.570796, 1.649399],accel_mss,speed_ms,0,blend_radius_m)
  movel([0.072873, -0.622675, -2.819228, -1.270485, 1.570796, 1.643669],accel_mss,speed_ms,0,blend_radius_m)
  movel([0.070007, -0.624773, -2.819042, -1.268573, 1.570796, 1.640803],accel_mss,speed_ms,0,blend_radius_m)
  speed_ms = 0.005
  movel([0.070007, -0.618828, -2.812252, -1.281309, 1.570796, 1.640803],accel_mss,speed_ms,0,blend_radius_m)
  speed_ms = 0.040
  movel([0.089300, -0.598858, -2.813943, -1.299588, 1.570796, 1.660097],accel_mss,speed_ms,0,blend_radius_m)
  speed_ms = 0.005
  movel([0.089300, -0.604471, -2.820769, -1.287149, 1.570796, 1.660097],accel_mss,speed_ms,0,blend_radius_m)
  speed_ms = 0.025
  movel([0.085848, -0.602247, -2.820948, -1.289194, 1.570796, 1.656644],accel_mss,speed_ms,0,blend_radius_m)
  movel([0.081583, -0.601122, -2.821038, -1.290229, 1.570796, 1.652379],accel_mss,speed_ms,0,blend_radius_m)
  movel([0.076593, -0.601161, -2.821035, -1.290193, 1.570796, 1.647389],accel_mss,speed_ms,0,blend_radius_m)
  movel([0.070948, -0.602405, -2.820935, -1.289049, 1.570796, 1.641744],accel_mss,speed_ms,0,blend_radius_m)
  movel([0.064745, -0.604900, -2.820734, -1.286755, 1.570796, 1.635541],accel_mss,speed_ms,0,blend_radius_m)
  movel([0.061464, -0.606623, -2.820593, -1.285173, 1.570796, 1.632260],accel_mss,speed_ms,0,blend_radius_m)
  movel([0.058084, -0.608666, -2.820425, -1.283297, 1.570796, 1.628881],accel_mss,speed_ms,0,blend_radius_m)
  movel([0.054609, -0.611039, -2.820228, -1.281123, 1.570796, 1.625405],accel_mss,speed_ms,0,blend_radius_m)
  movel([0.051053, -0.613741, -2.820000, -1.278647, 1.570796, 1.621849],accel_mss,speed_ms,0,blend_radius_m)
  movel([0.047438, -0.616765, -2.819743, -1.275881, 1.570796, 1.618234],accel_mss,speed_ms,0,blend_radius_m)
  movel([0.043773, -0.620117, -2.819453, -1.272820, 1.570796, 1.614569],accel_mss,speed_ms,0,blend_radius_m)
  speed_ms = 0.005
  movel([0.043773, -0.614246, -2.812654, -1.285489, 1.570796, 1.614569],accel_mss,speed_ms,0,blend_radius_m)
  speed_ms = 0.040
  movel([0.064233, -0.590185, -2.814629, -1.307575, 1.570796, 1.635029],accel_mss,speed_ms,0,blend_radius_m)
  speed_ms = 0.005
  movel([0.064233, -0.595651, -2.821468, -1.295270, 1.570796, 1.635029],accel_mss,speed_ms,0,blend_radius_m)
  speed_ms = 0.025
  movel([0.063094, -0.593144, -2.821662, -1.297583, 1.570796, 1.633890],accel_mss,speed_ms,0,blend_radius_m)
  movel([0.061364, -0.591307, -2.821802, -1.299280, 1.570796, 1.632160],accel_mss,speed_ms,0,blend_radius_m)
  movel([0.059073, -0.590179, -2.821887, -1.300323, 1.570796, 1.629869],accel_mss,speed_ms,0,blend_radius_m)
  movel([0.056266, -0.589792, -2.821917, -1.300680, 1.570796, 1.627062],accel_mss,speed_ms,0,blend_radius_m)
  movel([0.052290, -0.590281, -2.821880, -1.300228, 1.570796, 1.623086],accel_mss,speed_ms,0,blend_radius_m)
  movel([0.047869, -0.591585, -2.821781, -1.299023, 1.570796, 1.618665],accel_mss,speed_ms,0,blend_radius_m)
  movel([0.042312, -0.593872, -2.821606, -1.296911, 1.570796, 1.613109],accel_mss,speed_ms,0,blend_radius_m)
  movel([0.036448, -0.596965, -2.821366, -1.294058, 1.570796, 1.607244],accel_mss,speed_ms,0,blend_radius_m)
  movel([0.030360, -0.600886, -2.821057, -1.290446, 1.570796, 1.601157],accel_mss,speed_ms,0,blend_radius_m)
  movel([0.024131, -0.605669, -2.820671, -1.286048, 1.570796, 1.594927],accel_mss,speed_ms,0,blend_radius_m)
  movel([0.017873, -0.611324, -2.820204, -1.280861, 1.570796, 1.588669],accel_mss,speed_ms,0,blend_radius_m)
  movel([0.014803, -0.614432, -2.819942, -1.278015, 1.570796, 1.585600],accel_mss,speed_ms,0,blend_radius_m)
  movel([0.008947, -0.621082, -2.819368, -1.271939, 1.570796, 1.579743],accel_mss,speed_ms,0,blend_radius_m)
  movel([0.006216, -0.624566, -2.819061, -1.268762, 1.570796, 1.577013],accel_mss,speed_ms,0,blend_radius_m)
  movel([0.003666, -0.628123, -2.818742, -1.265524, 1.570796, 1.574462],accel_mss,speed_ms,0,blend_radius_m)
  movel([0.001318, -0.631730, -2.818413, -1.262245, 1.570796, 1.572114],accel_mss,speed_ms,0,blend_radius_m)
  speed_ms = 0.005
  movel([0.001318, -0.625674, -2.811635, -1.275080, 1.570796, 1.572114],accel_mss,speed_ms,0,blend_radius_m)
  speed_ms = 0.040
  movel([0.022676, -0.592973, -2.814412, -1.305004, 1.570796, 1.593472],accel_mss,speed_ms,0,blend_radius_m)
  speed_ms = 0.005
  movel([0.022676, -0.598486, -2.821247, -1.292656, 1.570796, 1.593472],accel_mss,speed_ms,0,blend_radius_m)
  speed_ms = 0.025
  movel([0.015376, -0.601915, -2.820974, -1.289499, 1.570796, 1.586173],accel_mss,speed_ms,0,blend_radius_m)
  movel([0.007626, -0.606364, -2.820614, -1.285411, 1.570796, 1.578423],accel_mss,speed_ms,0,blend_radius_m)
  movel([-0.000368, -0.611799, -2.820164, -1.280425, 1.570796, 1.570428],accel_mss,speed_ms,0,blend_radius_m)
  movel([-0.004391, -0.614867, -2.819905, -1.277617, 1.570796, 1.566405],accel_mss,speed_ms,0,blend_radius_m)
  movel([-0.008399, -0.618167, -2.819622, -1.274600, 1.570796, 1.562398],accel_mss,speed_ms,0,blend_radius_m)
  movel([-0.012357, -0.621683, -2.819316, -1.271390, 1.570796, 1.558439],accel_mss,speed_ms,0,blend_radius_m)
  movel([-0.016240, -0.625405, -2.818986, -1.267998, 1.570796, 1.554557],accel_mss,speed_ms,0,blend_radius_m)
  movel([-0.020025, -0.629332, -2.818632, -1.264425, 1.570796, 1.550771],accel_mss,speed_ms,0,blend_radius_m)
  movel([-0.023687, -0.633458, -2.818254, -1.260677, 1.570796, 1.547109],accel_mss,speed_ms,0,blend_radius_m)
  movel([-0.027206, -0.637773, -2.817851, -1.256765, 1.570796, 1.543591],accel_mss,speed_ms,0,blend_radius_m)
  movel([-0.030543, -0.642266, -2.817424, -1.252699, 1.570796, 1.540253],accel_mss,speed_ms,0,blend_radius_m)
  movel([-0.033686, -0.646932, -2.816971, -1.248486, 1.570796, 1.537111],accel_mss,speed_ms,0,blend_radius_m)
  movel([-0.036604, -0.651767, -2.816492, -1.244130, 1.570796, 1.534193],accel_mss,speed_ms,0,blend_radius_m)
  speed_ms = 0.005
  movel([-0.036604, -0.645397, -2.809752, -1.257240, 1.570796, 1.534193],accel_mss,speed_ms,0,blend_radius_m)
  speed_ms = 0.040
  movel([-0.022149, -0.613326, -2.812733, -1.286330, 1.570796, 1.548647],accel_mss,speed_ms,0,blend_radius_m)
  speed_ms = 0.005
  movel([-0.022149, -0.619181, -2.819534, -1.273674, 1.570796, 1.548647],accel_mss,speed_ms,0,blend_radius_m)
  speed_ms = 0.025
  movel([-0.025873, -0.621233, -2.819355, -1.271801, 1.570796, 1.544923],accel_mss,speed_ms,0,blend_radius_m)
  movel([-0.029708, -0.623683, -2.819139, -1.269567, 1.570796, 1.541089],accel_mss,speed_ms,0,blend_radius_m)
  movel([-0.033605, -0.626502, -2.818888, -1.266999, 1.570796, 1.537191],accel_mss,speed_ms,0,blend_radius_m)
  movel([-0.037532, -0.629649, -2.818603, -1.264136, 1.570796, 1.533264],accel_mss,speed_ms,0,blend_radius_m)
  movel([-0.041453, -0.633099, -2.818287, -1.261003, 1.570796, 1.529343],accel_mss,speed_ms,0,blend_radius_m)
  movel([-0.045324, -0.636813, -2.817941, -1.257635, 1.570796, 1.525473],accel_mss,speed_ms,0,blend_radius_m)
  movel([-0.049105, -0.640750, -2.817569, -1.254070, 1.570796, 1.521691],accel_mss,speed_ms,0,blend_radius_m)
  movel([-0.052772, -0.644891, -2.817170, -1.250328, 1.570796, 1.518024],accel_mss,speed_ms,0,blend_radius_m)
  movel([-0.056275, -0.649189, -2.816749, -1.246451, 1.570796, 1.514522],accel_mss,speed_ms,0,blend_radius_m)
  movel([-0.059585, -0.653597, -2.816309, -1.242483, 1.570796, 1.511211],accel_mss,speed_ms,0,blend_radius_m)
  movel([-0.062677, -0.658069, -2.815854, -1.238466, 1.570796, 1.508120],accel_mss,speed_ms,0,blend_radius_m)
  movel([-0.065528, -0.662569, -2.815388, -1.234432, 1.570796, 1.505269],accel_mss,speed_ms,0,blend_radius_m)
  movel([-0.068119, -0.667053, -2.814916, -1.230420, 1.570796, 1.502677],accel_mss,speed_ms,0,blend_radius_m)
  movel([-0.070432, -0.671494, -2.814439, -1.226456, 1.570796, 1.500365],accel_mss,speed_ms,0,blend_radius_m)
  movel([-0.072431, -0.675835, -2.813965, -1.222588, 1.570796, 1.498365],accel_mss,speed_ms,0,blend_radius_m)
  movel([-0.074111, -0.680050, -2.813498, -1.218841, 1.570796, 1.496685],accel_mss,speed_ms,0,blend_radius_m)
  speed_ms = 0.005
  movel([-0.074111, -0.673260, -2.806815, -1.232314, 1.570796, 1.496685],accel_mss,speed_ms,0,blend_radius_m)
  speed_ms = 0.040
  movel([-0.066858, -0.646255, -2.809666, -1.256467, 1.570796, 1.503938],accel_mss,speed_ms,0,blend_radius_m)
  speed_ms = 0.005
  movel([-0.066858, -0.652638, -2.816405, -1.243346, 1.570796, 1.503938],accel_mss,speed_ms,0,blend_radius_m)
  speed_ms = 0.025
  movel([-0.070442, -0.654850, -2.816182, -1.241356, 1.570796, 1.500354],accel_mss,speed_ms,0,blend_radius_m)
  movel([-0.074094, -0.657655, -2.815896, -1.238838, 1.570796, 1.496702],accel_mss,speed_ms,0,blend_radius_m)
  movel([-0.077748, -0.660951, -2.815557, -1.235881, 1.570796, 1.493049],accel_mss,speed_ms,0,blend_radius_m)
  movel([-0.081363, -0.664641, -2.815171, -1.232577, 1.570796, 1.489434],accel_mss,speed_ms,0,blend_radius_m)
  movel([-0.084887, -0.668634, -2.814747, -1.229008, 1.570796, 1.485909],accel_mss,speed_ms,0,blend_radius_m)
  movel([-0.088268, -0.672828, -2.814294, -1.225266, 1.570796, 1.482528],accel_mss,speed_ms,0,blend_radius_m)
  movel([-0.091469, -0.677133, -2.813822, -1.221434, 1.570796, 1.479327],accel_mss,speed_ms,0,blend_radius_m)
  movel([-0.094435, -0.681456, -2.813340, -1.217593, 1.570796, 1.476361],accel_mss,speed_ms,0,blend_radius_m)
  movel([-0.097268, -0.685917, -2.812834, -1.213638, 1.570796, 1.473529],accel_mss,speed_ms,0,blend_radius_m)
  movel([-0.099872, -0.690389, -2.812318, -1.209682, 1.570796, 1.470924],accel_mss,speed_ms,0,blend_radius_m)
  movel([-0.102209, -0.694820, -2.811799, -1.205770, 1.570796, 1.468587],accel_mss,speed_ms,0,blend_radius_m)
  movel([-0.104211, -0.699139, -2.811284, -1.201967, 1.570796, 1.466585],accel_mss,speed_ms,0,blend_radius_m)
  movel([-0.105837, -0.703282, -2.810782, -1.198325, 1.570796, 1.464959],accel_mss,speed_ms,0,blend_radius_m)
  movel([-0.107039, -0.707193, -2.810302, -1.194895, 1.570796, 1.463757],accel_mss,speed_ms,0,blend_radius_m)
  movel([-0.107755, -0.710804, -2.809852, -1.191733, 1.570796, 1.463041],accel_mss,speed_ms,0,blend_radius_m)
  movel([-0.107950, -0.714063, -2.809441, -1.188884, 1.570796, 1.462846],accel_mss,speed_ms,0,blend_radius_m)
  speed_ms = 0.005
  movel([-0.107950, -0.706799, -2.802836, -1.202754, 1.570796, 1.462846],accel_mss,speed_ms,0,blend_radius_m)
  speed_ms = 0.040
  movel([-0.110320, -0.689472, -2.804954, -1.217964, 1.570796, 1.460476],accel_mss,speed_ms,0,blend_radius_m)
  speed_ms = 0.005
  movel([-0.110320, -0.696496, -2.811600, -1.204293, 1.570796, 1.460476],accel_mss,speed_ms,0,blend_radius_m)
  speed_ms = 0.025
  movel([-0.115088, -0.701762, -2.810967, -1.199660, 1.570796, 1.455708],accel_mss,speed_ms,0,blend_radius_m)
  movel([-0.119860, -0.707643, -2.810246, -1.194500, 1.570796, 1.450936],accel_mss,speed_ms,0,blend_radius_m)
  movel([-0.124369, -0.713858, -2.809467, -1.189064, 1.570796, 1.446427],accel_mss,speed_ms,0,blend_radius_m)
  movel([-0.128353, -0.720131, -2.808663, -1.183594, 1.570796, 1.442443],accel_mss,speed_ms,0,blend_radius_m)
  movel([-0.131570, -0.726206, -2.807868, -1.178315, 1.570796, 1.439226],accel_mss,speed_ms,0,blend_radius_m)
  movel([-0.132817, -0.729095, -2.807484, -1.175811, 1.570796, 1.437979],accel_mss,speed_ms,0,blend_radius_m)
  movel([-0.133780, -0.731834, -2.807116, -1.173439, 1.570796, 1.437016],accel_mss,speed_ms,0,blend_radius_m)
  movel([-0.134435, -0.734408, -2.806767, -1.171214, 1.570796, 1.436361],accel_mss,speed_ms,0,blend_radius_m)
  movel([-0.134755, -0.736782, -2.806443, -1.169164, 1.570796, 1.436041],accel_mss,speed_ms,0,blend_radius_m)
  movel([-0.134702, -0.738917, -2.806149, -1.167323, 1.570796, 1.436094],accel_mss,speed_ms,0,blend_radius_m)
  movel([-0.134258, -0.740802, -2.805887, -1.165700, 1.570796, 1.436538],accel_mss,speed_ms,0,blend_radius_m)
  speed_ms = 0.005
  movel([-0.134258, -0.733191, -2.799348, -1.179850, 1.570796, 1.436538],accel_mss,speed_ms,0,blend_radius_m)
  speed_ms = 0.040
  movel([-0.143177, -0.732182, -2.799487, -1.180720, 1.570796, 1.427620],accel_mss,speed_ms,0,blend_radius_m)
  speed_ms = 0.005
  movel([-0.143177, -0.739780, -2.806029, -1.166579, 1.570796, 1.427620],accel_mss,speed_ms,0,blend_radius_m)
  speed_ms = 0.025
  movel([-0.148309, -0.748493, -2.804804, -1.159093, 1.570796, 1.422487],accel_mss,speed_ms,0,blend_radius_m)
  movel([-0.150599, -0.752852, -2.804177, -1.155360, 1.570796, 1.420197],accel_mss,speed_ms,0,blend_radius_m)
  movel([-0.152589, -0.757110, -2.803556, -1.151723, 1.570796, 1.418207],accel_mss,speed_ms,0,blend_radius_m)
  movel([-0.154194, -0.761204, -2.802951, -1.148234, 1.570796, 1.416602],accel_mss,speed_ms,0,blend_radius_m)
  movel([-0.155337, -0.765074, -2.802371, -1.144944, 1.570796, 1.415460],accel_mss,speed_ms,0,blend_radius_m)
  movel([-0.155927, -0.768645, -2.801830, -1.141914, 1.570796, 1.414869],accel_mss,speed_ms,0,blend_radius_m)
  movel([-0.155895, -0.771867, -2.801336, -1.139186, 1.570796, 1.414902],accel_mss,speed_ms,0,blend_radius_m)
  speed_ms = 0.005
  movel([-0.155895, -0.735669, -2.768871, -1.207849, 1.570796, 1.414902],accel_mss,speed_ms,0,blend_radius_m)
  speed_ms = 1.000
  movel([-0.155895, -0.735669, -2.768871, -1.207849, 1.570796, 1.414902],accel_mss,speed_ms,0,blend_radius_m)
  # Splitting Linear movement in 6 (instruction 3389: MoveL 3112)
  movel([-0.155895, -0.711776, -2.741501, -1.259111, 1.570796, 1.414902],accel_mss,speed_ms,0,blend_radius_m)
  movel([-0.155895, -0.692545, -2.713882, -1.305962, 1.570796, 1.414902],accel_mss,speed_ms,0,blend_radius_m)
  movel([-0.155895, -0.677214, -2.686036, -1.349139, 1.570796, 1.414902],accel_mss,speed_ms,0,blend_radius_m)
  movel([-0.155895, -0.665174, -2.657980, -1.389234, 1.570796, 1.414902],accel_mss,speed_ms,0,blend_radius_m)
  movel([-0.155895, -0.655937, -2.629727, -1.426724, 1.570796, 1.414902],accel_mss,speed_ms,0,blend_radius_m)
  movel([-0.155895, -0.649105, -2.601284, -1.462000, 1.570796, 1.414902],accel_mss,speed_ms,0,blend_radius_m)
  # End of main program
end

Machining1()
